// TIA Portal V20 export
TYPE "Keyence_Wert_lesen"
   STRUCT
      Read : Bool;   // Datensatzübertragung durchführen
      ID : HW_IO;   // Hardware-Kennung der Hardware-Baugruppe
      Index : DInt;   // Datensatznummer
      MLen : UInt;   // Maximale Länge der zu lesenden Datensatzinformation in Byte.
      Valid : Bool;   // Neuer Datensatz wurde empfangen und ist gültig.
      Busy : Bool;   // BUSY = 1: Der Lesevorgang ist noch nicht beendet.
      Error : Bool;   // ERROR = 1: Beim Lesevorgang trat ein Fehler auf.
      Status : DWord;   // Bausteinstatus bzw. Fehlerinformation.
      Len : UInt;   // Länge der gelesenen Datensatzinformation
      Record : DInt;   // Zielbereich für den gelesenen Datensatz.
   END_STRUCT;
END_TYPE
